// TIA Portal V20 export
Screen "Pop-up_SYSTEM_DIAGNOSTIC_LEGEND_Popup"  330x313
  ScreenItem "Background" at 0,0 size 330x313  Type=HmiRectangle
  ScreenItem "Text_Legend" at 1,1 size 328x25  Type=HmiTextBox
  ScreenItem "Text_DeviceInOperation" at 35,38 size 200x20  Type=HmiTextBox
  ScreenItem "Cancel Mode" at 239,1 size 90x61  Type=HmiButton
  ScreenItem "Graphic_DeviceInOperation" at 10,38 size 20x20  Type=HmiGraphicView
  ScreenItem "Graphic_DeviceCannotBeAccessed" at 10,61 size 20x20  Type=HmiGraphicView
  ScreenItem "Text_DeviceCannotBeAccessed" at 35,61 size 200x20  Type=HmiTextBox
  ScreenItem "Graphic_ErrorsInDevice" at 10,85 size 20x20  Type=HmiGraphicView
  ScreenItem "Text_ErrorsInDevice" at 35,85 size 285x20  Type=HmiTextBox
  ScreenItem "Graphic_DeviceDeactivated" at 10,107 size 20x20  Type=HmiGraphicView
  ScreenItem "Text_DeviceDeactivated" at 35,107 size 285x20  Type=HmiTextBox
  ScreenItem "Graphic_InputOutputDataNotAvailable" at 10,130 size 20x20  Type=HmiGraphicView
  ScreenItem "Text_InputOutputDataNotAvailable" at 35,130 size 285x20  Type=HmiTextBox
  ScreenItem "Graphic_MaintenanceRequired" at 10,153 size 20x20  Type=HmiGraphicView
  ScreenItem "Text_MaintenanceRequired" at 35,153 size 285x20  Type=HmiTextBox
  ScreenItem "Graphic_MaintenanceRecommended" at 10,176 size 20x20  Type=HmiGraphicView
  ScreenItem "Text_MaintenanceRecommended" at 35,176 size 285x20  Type=HmiTextBox
  ScreenItem "Text_SuperimposedSymbol" at 35,268 size 285x35  Type=HmiTextBox
  ScreenItem "Text_CurrentConfiguration" at 35,199 size 285x20  Type=HmiTextBox
  ScreenItem "Graphic_CurrentConfiguration" at 10,199 size 20x20  Type=HmiGraphicView
  ScreenItem "Graphic_SuperimposedSymbol" at 10,268 size 20x20  Type=HmiGraphicView
  ScreenItem "Text_StopEgUpdateBootOwnInitialization" at 35,222 size 285x20  Type=HmiTextBox
  ScreenItem "Text_Stop" at 35,245 size 285x20  Type=HmiTextBox
  ScreenItem "Graphic_StopEgUpdateBootOwnInitialization" at 10,222 size 20x20  Type=HmiGraphicView
  ScreenItem "Graphic_Stop" at 10,246 size 20x18  Type=HmiGraphicView
